FUNCTION_BLOCK FB_PERIPHERY_REF
VAR_INPUT

END_VAR
VAR_OUTPUT

END_VAR
VAR_IN_OUT

END_VAR
VAR

END_VAR

;

END_FUNCTION_BLOCK

(* stored: Version 1.1.0.1, ProductVersion 3.1.4024.15
   POU FB_PERIPHERY_REF: Id {ce294a97-136c-4ee4-920c-dda8f0bdd5e6}, SpecialFunc None *)
